(* IEC 61131-3 sources: trust-platform/examples/rust_first_cell/src/generated/trust, 2 files *)

(* ---- configuration.st ---- *)
(* GENERATED by trust-runtime from trust.toml - do not edit *)
CONFIGURATION CellRes
RESOURCE CellRes ON PLC
    TASK CellTask (INTERVAL := T#10ms, PRIORITY := 1);
    PROGRAM Cell WITH CellTask : PRESS_CELL;
END_RESOURCE
VAR_CONFIG
    Cell.start AT %IX0.0 : BOOL;
    Cell.part_present AT %IX0.1 : BOOL;
    Cell.clamp_closed AT %IX0.2 : BOOL;
    Cell.press_down AT %IX0.3 : BOOL;
    Cell.clamp AT %QX0.0 : BOOL;
    Cell.press AT %QX0.1 : BOOL;
    Cell.ready AT %QX0.2 : BOOL;
END_VAR
END_CONFIGURATION

(* ---- rust_pous.st ---- *)
(* GENERATED by trust-runtime from src/lib.rs - do not edit *)
TYPE
    PRESS_CELL_SEQ :
    STRUCT
        point : UINT;
        began : TIME;
        shape_a4638268 : BOOL;
    END_STRUCT;
END_TYPE

(* GENERATED by trust-runtime from src/lib.rs - do not edit *)
{attribute 'rust'}
PROGRAM PRESS_CELL
VAR_INPUT
    start : BOOL;
    part_present : BOOL;
    clamp_closed : BOOL;
    press_down : BOOL;
END_VAR
VAR_OUTPUT
    clamp : BOOL;
    press : BOOL;
    ready : BOOL;
    active_step : STRING[16];
    parts : UDINT;
END_VAR
VAR
    _seq : PRESS_CELL_SEQ;
END_VAR
END_PROGRAM
